Fanuc KAREL source: kt00475.KL

PROGRAM KT00475
%STACKSIZE=65535
%PRIORITY=65535
%NOLOCKGROUP
VAR
P1 : POSITION
P2 : POSITION
OUT : XYZWPR
BEGIN
-- UNRESOLVED_PC line 8 opcodes [49 49 60 7E 4A] marker_code=0
END KT00475
